Yaskawa INFORM job: VEGG2.JBI

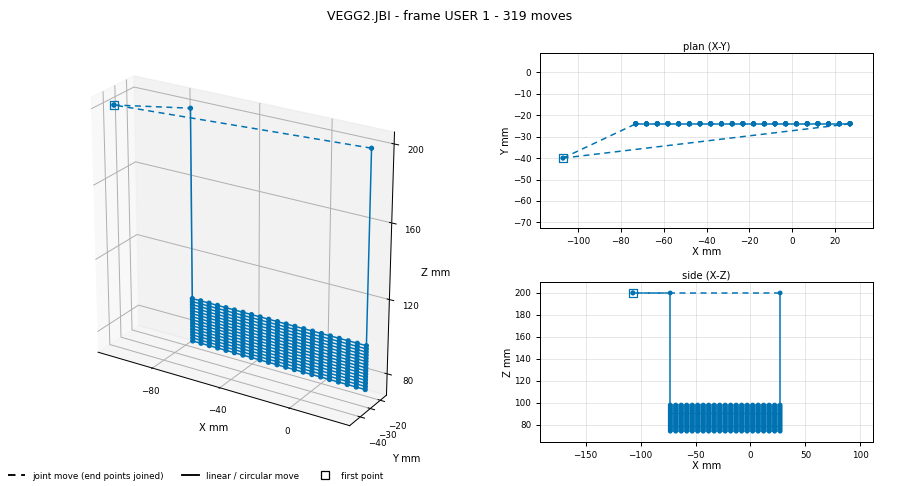
[picture p0: tool path of VEGG2.JBI in frame USER 1, 319 of 319 moves have a stored position in this frame; points joined in program order, loops and branches not executed]
/JOB
//NAME VEGG2
//POS
///NPOS 319,0,0,0,0,0
///USER 1
///TOOL 1
///POSTYPE USER
///RECTAN
///RCONF 1,0,0,0,0,0,0,0,0,0,0,0,0,0,0,0,0,0,0,0,0,0,0,0
C00000=-107.000,-40.000,200.000,0.0000,0.0000,-150.0000
C00001=-73.000,-24.000,200.000,0.0000,0.0000,-150.0000
C00002=-73.000,-24.000,74.200,0.0000,0.0000,-150.0000
C00003=-68.000,-24.000,74.200,0.0000,0.0000,-150.0000
C00004=-63.000,-24.000,74.200,0.0000,0.0000,-150.0000
C00005=-58.000,-24.000,74.200,0.0000,0.0000,-150.0000
C00006=-53.000,-24.000,74.200,0.0000,0.0000,-150.0000
C00007=-48.000,-24.000,74.200,0.0000,0.0000,-150.0000
C00008=-43.000,-24.000,74.200,0.0000,0.0000,-150.0000
C00009=-38.000,-24.000,74.200,0.0000,0.0000,-150.0000
C00010=-33.000,-24.000,74.200,0.0000,0.0000,-150.0000
C00011=-28.000,-24.000,74.200,0.0000,0.0000,-150.0000
C00012=-23.000,-24.000,74.200,0.0000,0.0000,-150.0000
C00013=-18.000,-24.000,74.200,0.0000,0.0000,-150.0000
C00014=-13.000,-24.000,74.200,0.0000,0.0000,-150.0000
C00015=-8.000,-24.000,74.200,0.0000,0.0000,-150.0000
C00016=-3.000,-24.000,74.200,0.0000,0.0000,-150.0000
C00017=2.000,-24.000,74.200,0.0000,0.0000,-150.0000
C00018=7.000,-24.000,74.200,0.0000,0.0000,-150.0000
C00019=12.000,-24.000,74.200,0.0000,0.0000,-150.0000
C00020=17.000,-24.000,74.200,0.0000,0.0000,-150.0000
C00021=22.000,-24.000,74.200,0.0000,0.0000,-150.0000
C00022=27.000,-24.000,74.200,0.0000,0.0000,-150.0000
C00023=27.000,-24.000,75.900,0.0000,0.0000,-150.0000
C00024=22.000,-24.000,75.900,0.0000,0.0000,-150.0000
C00025=17.000,-24.000,75.900,0.0000,0.0000,-150.0000
C00026=12.000,-24.000,75.900,0.0000,0.0000,-150.0000
C00027=7.000,-24.000,75.900,0.0000,0.0000,-150.0000
C00028=2.000,-24.000,75.900,0.0000,0.0000,-150.0000
C00029=-3.000,-24.000,75.900,0.0000,0.0000,-150.0000
C00030=-8.000,-24.000,75.900,0.0000,0.0000,-150.0000
C00031=-13.000,-24.000,75.900,0.0000,0.0000,-150.0000
C00032=-18.000,-24.000,75.900,0.0000,0.0000,-150.0000
C00033=-23.000,-24.000,75.900,0.0000,0.0000,-150.0000
C00034=-28.000,-24.000,75.900,0.0000,0.0000,-150.0000
C00035=-33.000,-24.000,75.900,0.0000,0.0000,-150.0000
C00036=-38.000,-24.000,75.900,0.0000,0.0000,-150.0000
C00037=-43.000,-24.000,75.900,0.0000,0.0000,-150.0000
C00038=-48.000,-24.000,75.900,0.0000,0.0000,-150.0000
C00039=-53.000,-24.000,75.900,0.0000,0.0000,-150.0000
C00040=-58.000,-24.000,75.900,0.0000,0.0000,-150.0000
C00041=-63.000,-24.000,75.900,0.0000,0.0000,-150.0000
C00042=-68.000,-24.000,75.900,0.0000,0.0000,-150.0000
C00043=-73.000,-24.000,75.900,0.0000,0.0000,-150.0000
C00044=-73.000,-24.000,77.600,0.0000,0.0000,-150.0000
C00045=-68.000,-24.000,77.600,0.0000,0.0000,-150.0000
C00046=-63.000,-24.000,77.600,0.0000,0.0000,-150.0000
C00047=-58.000,-24.000,77.600,0.0000,0.0000,-150.0000
C00048=-53.000,-24.000,77.600,0.0000,0.0000,-150.0000
C00049=-48.000,-24.000,77.600,0.0000,0.0000,-150.0000
C00050=-43.000,-24.000,77.600,0.0000,0.0000,-150.0000
C00051=-38.000,-24.000,77.600,0.0000,0.0000,-150.0000
C00052=-33.000,-24.000,77.600,0.0000,0.0000,-150.0000
C00053=-28.000,-24.000,77.600,0.0000,0.0000,-150.0000
C00054=-23.000,-24.000,77.600,0.0000,0.0000,-150.0000
C00055=-18.000,-24.000,77.600,0.0000,0.0000,-150.0000
C00056=-13.000,-24.000,77.600,0.0000,0.0000,-150.0000
C00057=-8.000,-24.000,77.600,0.0000,0.0000,-150.0000
C00058=-3.000,-24.000,77.600,0.0000,0.0000,-150.0000
C00059=2.000,-24.000,77.600,0.0000,0.0000,-150.0000
C00060=7.000,-24.000,77.600,0.0000,0.0000,-150.0000
C00061=12.000,-24.000,77.600,0.0000,0.0000,-150.0000
C00062=17.000,-24.000,77.600,0.0000,0.0000,-150.0000
C00063=22.000,-24.000,77.600,0.0000,0.0000,-150.0000
C00064=27.000,-24.000,77.600,0.0000,0.0000,-150.0000
C00065=27.000,-24.000,79.300,0.0000,0.0000,-150.0000
C00066=22.000,-24.000,79.300,0.0000,0.0000,-150.0000
C00067=17.000,-24.000,79.300,0.0000,0.0000,-150.0000
C00068=12.000,-24.000,79.300,0.0000,0.0000,-150.0000
C00069=7.000,-24.000,79.300,0.0000,0.0000,-150.0000
C00070=2.000,-24.000,79.300,0.0000,0.0000,-150.0000
C00071=-3.000,-24.000,79.300,0.0000,0.0000,-150.0000
C00072=-8.000,-24.000,79.300,0.0000,0.0000,-150.0000
C00073=-13.000,-24.000,79.300,0.0000,0.0000,-150.0000
C00074=-18.000,-24.000,79.300,0.0000,0.0000,-150.0000
C00075=-23.000,-24.000,79.300,0.0000,0.0000,-150.0000
C00076=-28.000,-24.000,79.300,0.0000,0.0000,-150.0000
C00077=-33.000,-24.000,79.300,0.0000,0.0000,-150.0000
C00078=-38.000,-24.000,79.300,0.0000,0.0000,-150.0000
C00079=-43.000,-24.000,79.300,0.0000,0.0000,-150.0000
C00080=-48.000,-24.000,79.300,0.0000,0.0000,-150.0000
C00081=-53.000,-24.000,79.300,0.0000,0.0000,-150.0000
C00082=-58.000,-24.000,79.300,0.0000,0.0000,-150.0000
C00083=-63.000,-24.000,79.300,0.0000,0.0000,-150.0000
C00084=-68.000,-24.000,79.300,0.0000,0.0000,-150.0000
C00085=-73.000,-24.000,79.300,0.0000,0.0000,-150.0000
C00086=-73.000,-24.000,81.000,0.0000,0.0000,-150.0000
C00087=-68.000,-24.000,81.000,0.0000,0.0000,-150.0000
C00088=-63.000,-24.000,81.000,0.0000,0.0000,-150.0000
C00089=-58.000,-24.000,81.000,0.0000,0.0000,-150.0000
C00090=-53.000,-24.000,81.000,0.0000,0.0000,-150.0000
C00091=-48.000,-24.000,81.000,0.0000,0.0000,-150.0000
C00092=-43.000,-24.000,81.000,0.0000,0.0000,-150.0000
C00093=-38.000,-24.000,81.000,0.0000,0.0000,-150.0000
C00094=-33.000,-24.000,81.000,0.0000,0.0000,-150.0000
C00095=-28.000,-24.000,81.000,0.0000,0.0000,-150.0000
C00096=-23.000,-24.000,81.000,0.0000,0.0000,-150.0000
C00097=-18.000,-24.000,81.000,0.0000,0.0000,-150.0000
C00098=-13.000,-24.000,81.000,0.0000,0.0000,-150.0000
C00099=-8.000,-24.000,81.000,0.0000,0.0000,-150.0000
C00100=-3.000,-24.000,81.000,0.0000,0.0000,-150.0000
C00101=2.000,-24.000,81.000,0.0000,0.0000,-150.0000
C00102=7.000,-24.000,81.000,0.0000,0.0000,-150.0000
C00103=12.000,-24.000,81.000,0.0000,0.0000,-150.0000
C00104=17.000,-24.000,81.000,0.0000,0.0000,-150.0000
C00105=22.000,-24.000,81.000,0.0000,0.0000,-150.0000
C00106=27.000,-24.000,81.000,0.0000,0.0000,-150.0000
C00107=27.000,-24.000,82.700,0.0000,0.0000,-150.0000
C00108=22.000,-24.000,82.700,0.0000,0.0000,-150.0000
C00109=17.000,-24.000,82.700,0.0000,0.0000,-150.0000
C00110=12.000,-24.000,82.700,0.0000,0.0000,-150.0000
C00111=7.000,-24.000,82.700,0.0000,0.0000,-150.0000
C00112=2.000,-24.000,82.700,0.0000,0.0000,-150.0000
C00113=-3.000,-24.000,82.700,0.0000,0.0000,-150.0000
C00114=-8.000,-24.000,82.700,0.0000,0.0000,-150.0000
C00115=-13.000,-24.000,82.700,0.0000,0.0000,-150.0000
C00116=-18.000,-24.000,82.700,0.0000,0.0000,-150.0000
C00117=-23.000,-24.000,82.700,0.0000,0.0000,-150.0000
C00118=-28.000,-24.000,82.700,0.0000,0.0000,-150.0000
C00119=-33.000,-24.000,82.700,0.0000,0.0000,-150.0000
C00120=-38.000,-24.000,82.700,0.0000,0.0000,-150.0000
C00121=-43.000,-24.000,82.700,0.0000,0.0000,-150.0000
C00122=-48.000,-24.000,82.700,0.0000,0.0000,-150.0000
C00123=-53.000,-24.000,82.700,0.0000,0.0000,-150.0000
C00124=-58.000,-24.000,82.700,0.0000,0.0000,-150.0000
C00125=-63.000,-24.000,82.700,0.0000,0.0000,-150.0000
C00126=-68.000,-24.000,82.700,0.0000,0.0000,-150.0000
C00127=-73.000,-24.000,82.700,0.0000,0.0000,-150.0000
C00128=-73.000,-24.000,84.400,0.0000,0.0000,-150.0000
C00129=-68.000,-24.000,84.400,0.0000,0.0000,-150.0000
C00130=-63.000,-24.000,84.400,0.0000,0.0000,-150.0000
C00131=-58.000,-24.000,84.400,0.0000,0.0000,-150.0000
C00132=-53.000,-24.000,84.400,0.0000,0.0000,-150.0000
C00133=-48.000,-24.000,84.400,0.0000,0.0000,-150.0000
C00134=-43.000,-24.000,84.400,0.0000,0.0000,-150.0000
C00135=-38.000,-24.000,84.400,0.0000,0.0000,-150.0000
C00136=-33.000,-24.000,84.400,0.0000,0.0000,-150.0000
C00137=-28.000,-24.000,84.400,0.0000,0.0000,-150.0000
C00138=-23.000,-24.000,84.400,0.0000,0.0000,-150.0000
C00139=-18.000,-24.000,84.400,0.0000,0.0000,-150.0000
C00140=-13.000,-24.000,84.400,0.0000,0.0000,-150.0000
C00141=-8.000,-24.000,84.400,0.0000,0.0000,-150.0000
C00142=-3.000,-24.000,84.400,0.0000,0.0000,-150.0000
C00143=2.000,-24.000,84.400,0.0000,0.0000,-150.0000
C00144=7.000,-24.000,84.400,0.0000,0.0000,-150.0000
C00145=12.000,-24.000,84.400,0.0000,0.0000,-150.0000
C00146=17.000,-24.000,84.400,0.0000,0.0000,-150.0000
C00147=22.000,-24.000,84.400,0.0000,0.0000,-150.0000
C00148=27.000,-24.000,84.400,0.0000,0.0000,-150.0000
C00149=27.000,-24.000,86.100,0.0000,0.0000,-150.0000
C00150=22.000,-24.000,86.100,0.0000,0.0000,-150.0000
C00151=17.000,-24.000,86.100,0.0000,0.0000,-150.0000
C00152=12.000,-24.000,86.100,0.0000,0.0000,-150.0000
C00153=7.000,-24.000,86.100,0.0000,0.0000,-150.0000
C00154=2.000,-24.000,86.100,0.0000,0.0000,-150.0000
C00155=-3.000,-24.000,86.100,0.0000,0.0000,-150.0000
C00156=-8.000,-24.000,86.100,0.0000,0.0000,-150.0000
C00157=-13.000,-24.000,86.100,0.0000,0.0000,-150.0000
C00158=-18.000,-24.000,86.100,0.0000,0.0000,-150.0000
C00159=-23.000,-24.000,86.100,0.0000,0.0000,-150.0000
C00160=-28.000,-24.000,86.100,0.0000,0.0000,-150.0000
C00161=-33.000,-24.000,86.100,0.0000,0.0000,-150.0000
C00162=-38.000,-24.000,86.100,0.0000,0.0000,-150.0000
C00163=-43.000,-24.000,86.100,0.0000,0.0000,-150.0000
C00164=-48.000,-24.000,86.100,0.0000,0.0000,-150.0000
C00165=-53.000,-24.000,86.100,0.0000,0.0000,-150.0000
C00166=-58.000,-24.000,86.100,0.0000,0.0000,-150.0000
C00167=-63.000,-24.000,86.100,0.0000,0.0000,-150.0000
C00168=-68.000,-24.000,86.100,0.0000,0.0000,-150.0000
C00169=-73.000,-24.000,86.100,0.0000,0.0000,-150.0000
C00170=-73.000,-24.000,87.800,0.0000,0.0000,-150.0000
C00171=-68.000,-24.000,87.800,0.0000,0.0000,-150.0000
C00172=-63.000,-24.000,87.800,0.0000,0.0000,-150.0000
C00173=-58.000,-24.000,87.800,0.0000,0.0000,-150.0000
C00174=-53.000,-24.000,87.800,0.0000,0.0000,-150.0000
C00175=-48.000,-24.000,87.800,0.0000,0.0000,-150.0000
C00176=-43.000,-24.000,87.800,0.0000,0.0000,-150.0000
C00177=-38.000,-24.000,87.800,0.0000,0.0000,-150.0000
C00178=-33.000,-24.000,87.800,0.0000,0.0000,-150.0000
C00179=-28.000,-24.000,87.800,0.0000,0.0000,-150.0000
C00180=-23.000,-24.000,87.800,0.0000,0.0000,-150.0000
C00181=-18.000,-24.000,87.800,0.0000,0.0000,-150.0000
C00182=-13.000,-24.000,87.800,0.0000,0.0000,-150.0000
C00183=-8.000,-24.000,87.800,0.0000,0.0000,-150.0000
C00184=-3.000,-24.000,87.800,0.0000,0.0000,-150.0000
C00185=2.000,-24.000,87.800,0.0000,0.0000,-150.0000
C00186=7.000,-24.000,87.800,0.0000,0.0000,-150.0000
C00187=12.000,-24.000,87.800,0.0000,0.0000,-150.0000
C00188=17.000,-24.000,87.800,0.0000,0.0000,-150.0000
C00189=22.000,-24.000,87.800,0.0000,0.0000,-150.0000
C00190=27.000,-24.000,87.800,0.0000,0.0000,-150.0000
C00191=27.000,-24.000,89.500,0.0000,0.0000,-150.0000
C00192=22.000,-24.000,89.500,0.0000,0.0000,-150.0000
C00193=17.000,-24.000,89.500,0.0000,0.0000,-150.0000
C00194=12.000,-24.000,89.500,0.0000,0.0000,-150.0000
C00195=7.000,-24.000,89.500,0.0000,0.0000,-150.0000
C00196=2.000,-24.000,89.500,0.0000,0.0000,-150.0000
C00197=-3.000,-24.000,89.500,0.0000,0.0000,-150.0000
C00198=-8.000,-24.000,89.500,0.0000,0.0000,-150.0000
C00199=-13.000,-24.000,89.500,0.0000,0.0000,-150.0000
C00200=-18.000,-24.000,89.500,0.0000,0.0000,-150.0000
C00201=-23.000,-24.000,89.500,0.0000,0.0000,-150.0000
C00202=-28.000,-24.000,89.500,0.0000,0.0000,-150.0000
C00203=-33.000,-24.000,89.500,0.0000,0.0000,-150.0000
C00204=-38.000,-24.000,89.500,0.0000,0.0000,-150.0000
C00205=-43.000,-24.000,89.500,0.0000,0.0000,-150.0000
C00206=-48.000,-24.000,89.500,0.0000,0.0000,-150.0000
C00207=-53.000,-24.000,89.500,0.0000,0.0000,-150.0000
C00208=-58.000,-24.000,89.500,0.0000,0.0000,-150.0000
C00209=-63.000,-24.000,89.500,0.0000,0.0000,-150.0000
C00210=-68.000,-24.000,89.500,0.0000,0.0000,-150.0000
C00211=-73.000,-24.000,89.500,0.0000,0.0000,-150.0000
C00212=-73.000,-24.000,91.200,0.0000,0.0000,-150.0000
C00213=-68.000,-24.000,91.200,0.0000,0.0000,-150.0000
C00214=-63.000,-24.000,91.200,0.0000,0.0000,-150.0000
C00215=-58.000,-24.000,91.200,0.0000,0.0000,-150.0000
C00216=-53.000,-24.000,91.200,0.0000,0.0000,-150.0000
C00217=-48.000,-24.000,91.200,0.0000,0.0000,-150.0000
C00218=-43.000,-24.000,91.200,0.0000,0.0000,-150.0000
C00219=-38.000,-24.000,91.200,0.0000,0.0000,-150.0000
C00220=-33.000,-24.000,91.200,0.0000,0.0000,-150.0000
C00221=-28.000,-24.000,91.200,0.0000,0.0000,-150.0000
C00222=-23.000,-24.000,91.200,0.0000,0.0000,-150.0000
C00223=-18.000,-24.000,91.200,0.0000,0.0000,-150.0000
C00224=-13.000,-24.000,91.200,0.0000,0.0000,-150.0000
C00225=-8.000,-24.000,91.200,0.0000,0.0000,-150.0000
C00226=-3.000,-24.000,91.200,0.0000,0.0000,-150.0000
C00227=2.000,-24.000,91.200,0.0000,0.0000,-150.0000
C00228=7.000,-24.000,91.200,0.0000,0.0000,-150.0000
C00229=12.000,-24.000,91.200,0.0000,0.0000,-150.0000
C00230=17.000,-24.000,91.200,0.0000,0.0000,-150.0000
C00231=22.000,-24.000,91.200,0.0000,0.0000,-150.0000
C00232=27.000,-24.000,91.200,0.0000,0.0000,-150.0000
C00233=27.000,-24.000,92.900,0.0000,0.0000,-150.0000
C00234=22.000,-24.000,92.900,0.0000,0.0000,-150.0000
C00235=17.000,-24.000,92.900,0.0000,0.0000,-150.0000
C00236=12.000,-24.000,92.900,0.0000,0.0000,-150.0000
C00237=7.000,-24.000,92.900,0.0000,0.0000,-150.0000
C00238=2.000,-24.000,92.900,0.0000,0.0000,-150.0000
C00239=-3.000,-24.000,92.900,0.0000,0.0000,-150.0000
C00240=-8.000,-24.000,92.900,0.0000,0.0000,-150.0000
C00241=-13.000,-24.000,92.900,0.0000,0.0000,-150.0000
C00242=-18.000,-24.000,92.900,0.0000,0.0000,-150.0000
C00243=-23.000,-24.000,92.900,0.0000,0.0000,-150.0000
C00244=-28.000,-24.000,92.900,0.0000,0.0000,-150.0000
C00245=-33.000,-24.000,92.900,0.0000,0.0000,-150.0000
C00246=-38.000,-24.000,92.900,0.0000,0.0000,-150.0000
C00247=-43.000,-24.000,92.900,0.0000,0.0000,-150.0000
C00248=-48.000,-24.000,92.900,0.0000,0.0000,-150.0000
C00249=-53.000,-24.000,92.900,0.0000,0.0000,-150.0000
C00250=-58.000,-24.000,92.900,0.0000,0.0000,-150.0000
C00251=-63.000,-24.000,92.900,0.0000,0.0000,-150.0000
C00252=-68.000,-24.000,92.900,0.0000,0.0000,-150.0000
C00253=-73.000,-24.000,92.900,0.0000,0.0000,-150.0000
C00254=-73.000,-24.000,94.600,0.0000,0.0000,-150.0000
C00255=-68.000,-24.000,94.600,0.0000,0.0000,-150.0000
C00256=-63.000,-24.000,94.600,0.0000,0.0000,-150.0000
C00257=-58.000,-24.000,94.600,0.0000,0.0000,-150.0000
C00258=-53.000,-24.000,94.600,0.0000,0.0000,-150.0000
C00259=-48.000,-24.000,94.600,0.0000,0.0000,-150.0000
C00260=-43.000,-24.000,94.600,0.0000,0.0000,-150.0000
C00261=-38.000,-24.000,94.600,0.0000,0.0000,-150.0000
C00262=-33.000,-24.000,94.600,0.0000,0.0000,-150.0000
C00263=-28.000,-24.000,94.600,0.0000,0.0000,-150.0000
C00264=-23.000,-24.000,94.600,0.0000,0.0000,-150.0000
C00265=-18.000,-24.000,94.600,0.0000,0.0000,-150.0000
C00266=-13.000,-24.000,94.600,0.0000,0.0000,-150.0000
C00267=-8.000,-24.000,94.600,0.0000,0.0000,-150.0000
C00268=-3.000,-24.000,94.600,0.0000,0.0000,-150.0000
C00269=2.000,-24.000,94.600,0.0000,0.0000,-150.0000
C00270=7.000,-24.000,94.600,0.0000,0.0000,-150.0000
C00271=12.000,-24.000,94.600,0.0000,0.0000,-150.0000
C00272=17.000,-24.000,94.600,0.0000,0.0000,-150.0000
C00273=22.000,-24.000,94.600,0.0000,0.0000,-150.0000
C00274=27.000,-24.000,94.600,0.0000,0.0000,-150.0000
C00275=27.000,-24.000,96.300,0.0000,0.0000,-150.0000
C00276=22.000,-24.000,96.300,0.0000,0.0000,-150.0000
C00277=17.000,-24.000,96.300,0.0000,0.0000,-150.0000
C00278=12.000,-24.000,96.300,0.0000,0.0000,-150.0000
C00279=7.000,-24.000,96.300,0.0000,0.0000,-150.0000
C00280=2.000,-24.000,96.300,0.0000,0.0000,-150.0000
C00281=-3.000,-24.000,96.300,0.0000,0.0000,-150.0000
C00282=-8.000,-24.000,96.300,0.0000,0.0000,-150.0000
C00283=-13.000,-24.000,96.300,0.0000,0.0000,-150.0000
C00284=-18.000,-24.000,96.300,0.0000,0.0000,-150.0000
C00285=-23.000,-24.000,96.300,0.0000,0.0000,-150.0000
C00286=-28.000,-24.000,96.300,0.0000,0.0000,-150.0000
C00287=-33.000,-24.000,96.300,0.0000,0.0000,-150.0000
C00288=-38.000,-24.000,96.300,0.0000,0.0000,-150.0000
C00289=-43.000,-24.000,96.300,0.0000,0.0000,-150.0000
C00290=-48.000,-24.000,96.300,0.0000,0.0000,-150.0000
C00291=-53.000,-24.000,96.300,0.0000,0.0000,-150.0000
C00292=-58.000,-24.000,96.300,0.0000,0.0000,-150.0000
C00293=-63.000,-24.000,96.300,0.0000,0.0000,-150.0000
C00294=-68.000,-24.000,96.300,0.0000,0.0000,-150.0000
C00295=-73.000,-24.000,96.300,0.0000,0.0000,-150.0000
C00296=-73.000,-24.000,98.000,0.0000,0.0000,-150.0000
C00297=-68.000,-24.000,98.000,0.0000,0.0000,-150.0000
C00298=-63.000,-24.000,98.000,0.0000,0.0000,-150.0000
C00299=-58.000,-24.000,98.000,0.0000,0.0000,-150.0000
C00300=-53.000,-24.000,98.000,0.0000,0.0000,-150.0000
C00301=-48.000,-24.000,98.000,0.0000,0.0000,-150.0000
C00302=-43.000,-24.000,98.000,0.0000,0.0000,-150.0000
C00303=-38.000,-24.000,98.000,0.0000,0.0000,-150.0000
C00304=-33.000,-24.000,98.000,0.0000,0.0000,-150.0000
C00305=-28.000,-24.000,98.000,0.0000,0.0000,-150.0000
C00306=-23.000,-24.000,98.000,0.0000,0.0000,-150.0000
C00307=-18.000,-24.000,98.000,0.0000,0.0000,-150.0000
C00308=-13.000,-24.000,98.000,0.0000,0.0000,-150.0000
C00309=-8.000,-24.000,98.000,0.0000,0.0000,-150.0000
C00310=-3.000,-24.000,98.000,0.0000,0.0000,-150.0000
C00311=2.000,-24.000,98.000,0.0000,0.0000,-150.0000
C00312=7.000,-24.000,98.000,0.0000,0.0000,-150.0000
C00313=12.000,-24.000,98.000,0.0000,0.0000,-150.0000
C00314=17.000,-24.000,98.000,0.0000,0.0000,-150.0000
C00315=22.000,-24.000,98.000,0.0000,0.0000,-150.0000
C00316=27.000,-24.000,98.000,0.0000,0.0000,-150.0000
C00317=27.000,-24.000,200.000,0.0000,0.0000,-150.0000
C00318=-107.000,-40.000,200.000,0.0000,0.0000,-150.0000
//INST
///DATE 2026/11/20 16:20
///ATTR SC,RW,RJ
////FRAME USER 1
///GROUP1 RB1
NOP
MOVJ C00000 VJ=0.78
MOVJ C00001 VJ=0.78
MOVL C00002 V=7.0 ACC=20 DEC=20
*LAG1
MACRO1 MJ#(0) ARGF1
ARCON
MOVL C00003 V=7.0 ACC=20 DEC=20
MOVL C00004 V=7.0 ACC=20 DEC=20
MOVL C00005 V=7.0 ACC=20 DEC=20
MOVL C00006 V=7.0 ACC=20 DEC=20
MOVL C00007 V=7.0 ACC=20 DEC=20
MOVL C00008 V=7.0 ACC=20 DEC=20
MOVL C00009 V=7.0 ACC=20 DEC=20
MOVL C00010 V=7.0 ACC=20 DEC=20
MOVL C00011 V=7.0 ACC=20 DEC=20
MOVL C00012 V=7.0 ACC=20 DEC=20
MOVL C00013 V=7.0 ACC=20 DEC=20
MOVL C00014 V=7.0 ACC=20 DEC=20
MOVL C00015 V=7.0 ACC=20 DEC=20
MOVL C00016 V=7.0 ACC=20 DEC=20
MOVL C00017 V=7.0 ACC=20 DEC=20
MOVL C00018 V=7.0 ACC=20 DEC=20
MOVL C00019 V=7.0 ACC=20 DEC=20
MOVL C00020 V=7.0 ACC=20 DEC=20
MOVL C00021 V=7.0 ACC=20 DEC=20
MOVL C00022 V=7.0 ACC=20 DEC=20
ARCOF
TIMER T=30
*LAG2
MOVL C00023 V=7.0 ACC=20 DEC=20
MACRO1 MJ#(0) ARGF2
ARCON
MOVL C00024 V=7.0 ACC=20 DEC=20
MOVL C00025 V=7.0 ACC=20 DEC=20
MOVL C00026 V=7.0 ACC=20 DEC=20
MOVL C00027 V=7.0 ACC=20 DEC=20
MOVL C00028 V=7.0 ACC=20 DEC=20
MOVL C00029 V=7.0 ACC=20 DEC=20
MOVL C00030 V=7.0 ACC=20 DEC=20
MOVL C00031 V=7.0 ACC=20 DEC=20
MOVL C00032 V=7.0 ACC=20 DEC=20
MOVL C00033 V=7.0 ACC=20 DEC=20
MOVL C00034 V=7.0 ACC=20 DEC=20
MOVL C00035 V=7.0 ACC=20 DEC=20
MOVL C00036 V=7.0 ACC=20 DEC=20
MOVL C00037 V=7.0 ACC=20 DEC=20
MOVL C00038 V=7.0 ACC=20 DEC=20
MOVL C00039 V=7.0 ACC=20 DEC=20
MOVL C00040 V=7.0 ACC=20 DEC=20
MOVL C00041 V=7.0 ACC=20 DEC=20
MOVL C00042 V=7.0 ACC=20 DEC=20
MOVL C00043 V=7.0 ACC=20 DEC=20
ARCOF
TIMER T=30
*LAG3
MOVL C00044 V=7.0 ACC=20 DEC=20
MACRO1 MJ#(0) ARGF2
ARCON
MOVL C00045 V=7.0 ACC=20 DEC=20
MOVL C00046 V=7.0 ACC=20 DEC=20
MOVL C00047 V=7.0 ACC=20 DEC=20
MOVL C00048 V=7.0 ACC=20 DEC=20
MOVL C00049 V=7.0 ACC=20 DEC=20
MOVL C00050 V=7.0 ACC=20 DEC=20
MOVL C00051 V=7.0 ACC=20 DEC=20
MOVL C00052 V=7.0 ACC=20 DEC=20
MOVL C00053 V=7.0 ACC=20 DEC=20
MOVL C00054 V=7.0 ACC=20 DEC=20
MOVL C00055 V=7.0 ACC=20 DEC=20
MOVL C00056 V=7.0 ACC=20 DEC=20
MOVL C00057 V=7.0 ACC=20 DEC=20
MOVL C00058 V=7.0 ACC=20 DEC=20
MOVL C00059 V=7.0 ACC=20 DEC=20
MOVL C00060 V=7.0 ACC=20 DEC=20
MOVL C00061 V=7.0 ACC=20 DEC=20
MOVL C00062 V=7.0 ACC=20 DEC=20
MOVL C00063 V=7.0 ACC=20 DEC=20
MOVL C00064 V=7.0 ACC=20 DEC=20
ARCOF
TIMER T=30
*LAG4
MOVL C00065 V=7.0 ACC=20 DEC=20
MACRO1 MJ#(0) ARGF2
ARCON
MOVL C00066 V=7.0 ACC=20 DEC=20
MOVL C00067 V=7.0 ACC=20 DEC=20
MOVL C00068 V=7.0 ACC=20 DEC=20
MOVL C00069 V=7.0 ACC=20 DEC=20
MOVL C00070 V=7.0 ACC=20 DEC=20
MOVL C00071 V=7.0 ACC=20 DEC=20
MOVL C00072 V=7.0 ACC=20 DEC=20
MOVL C00073 V=7.0 ACC=20 DEC=20
MOVL C00074 V=7.0 ACC=20 DEC=20
MOVL C00075 V=7.0 ACC=20 DEC=20
MOVL C00076 V=7.0 ACC=20 DEC=20
MOVL C00077 V=7.0 ACC=20 DEC=20
MOVL C00078 V=7.0 ACC=20 DEC=20
MOVL C00079 V=7.0 ACC=20 DEC=20
MOVL C00080 V=7.0 ACC=20 DEC=20
MOVL C00081 V=7.0 ACC=20 DEC=20
MOVL C00082 V=7.0 ACC=20 DEC=20
MOVL C00083 V=7.0 ACC=20 DEC=20
MOVL C00084 V=7.0 ACC=20 DEC=20
MOVL C00085 V=7.0 ACC=20 DEC=20
ARCOF
TIMER T=30
*LAG5
MOVL C00086 V=7.0 ACC=20 DEC=20
MACRO1 MJ#(0) ARGF2
ARCON
MOVL C00087 V=7.0 ACC=20 DEC=20
MOVL C00088 V=7.0 ACC=20 DEC=20
MOVL C00089 V=7.0 ACC=20 DEC=20
MOVL C00090 V=7.0 ACC=20 DEC=20
MOVL C00091 V=7.0 ACC=20 DEC=20
MOVL C00092 V=7.0 ACC=20 DEC=20
MOVL C00093 V=7.0 ACC=20 DEC=20
MOVL C00094 V=7.0 ACC=20 DEC=20
MOVL C00095 V=7.0 ACC=20 DEC=20
MOVL C00096 V=7.0 ACC=20 DEC=20
MOVL C00097 V=7.0 ACC=20 DEC=20
MOVL C00098 V=7.0 ACC=20 DEC=20
MOVL C00099 V=7.0 ACC=20 DEC=20
MOVL C00100 V=7.0 ACC=20 DEC=20
MOVL C00101 V=7.0 ACC=20 DEC=20
MOVL C00102 V=7.0 ACC=20 DEC=20
MOVL C00103 V=7.0 ACC=20 DEC=20
MOVL C00104 V=7.0 ACC=20 DEC=20
MOVL C00105 V=7.0 ACC=20 DEC=20
MOVL C00106 V=7.0 ACC=20 DEC=20
ARCOF
TIMER T=30
*LAG6
MOVL C00107 V=7.0 ACC=20 DEC=20
MACRO1 MJ#(0) ARGF2
ARCON
MOVL C00108 V=7.0 ACC=20 DEC=20
MOVL C00109 V=7.0 ACC=20 DEC=20
MOVL C00110 V=7.0 ACC=20 DEC=20
MOVL C00111 V=7.0 ACC=20 DEC=20
MOVL C00112 V=7.0 ACC=20 DEC=20
MOVL C00113 V=7.0 ACC=20 DEC=20
MOVL C00114 V=7.0 ACC=20 DEC=20
MOVL C00115 V=7.0 ACC=20 DEC=20
MOVL C00116 V=7.0 ACC=20 DEC=20
MOVL C00117 V=7.0 ACC=20 DEC=20
MOVL C00118 V=7.0 ACC=20 DEC=20
MOVL C00119 V=7.0 ACC=20 DEC=20
MOVL C00120 V=7.0 ACC=20 DEC=20
MOVL C00121 V=7.0 ACC=20 DEC=20
MOVL C00122 V=7.0 ACC=20 DEC=20
MOVL C00123 V=7.0 ACC=20 DEC=20
MOVL C00124 V=7.0 ACC=20 DEC=20
MOVL C00125 V=7.0 ACC=20 DEC=20
MOVL C00126 V=7.0 ACC=20 DEC=20
MOVL C00127 V=7.0 ACC=20 DEC=20
ARCOF
TIMER T=30
*LAG7
MOVL C00128 V=7.0 ACC=20 DEC=20
MACRO1 MJ#(0) ARGF2
ARCON
MOVL C00129 V=7.0 ACC=20 DEC=20
MOVL C00130 V=7.0 ACC=20 DEC=20
MOVL C00131 V=7.0 ACC=20 DEC=20
MOVL C00132 V=7.0 ACC=20 DEC=20
MOVL C00133 V=7.0 ACC=20 DEC=20
MOVL C00134 V=7.0 ACC=20 DEC=20
MOVL C00135 V=7.0 ACC=20 DEC=20
MOVL C00136 V=7.0 ACC=20 DEC=20
MOVL C00137 V=7.0 ACC=20 DEC=20
MOVL C00138 V=7.0 ACC=20 DEC=20
MOVL C00139 V=7.0 ACC=20 DEC=20
MOVL C00140 V=7.0 ACC=20 DEC=20
MOVL C00141 V=7.0 ACC=20 DEC=20
MOVL C00142 V=7.0 ACC=20 DEC=20
MOVL C00143 V=7.0 ACC=20 DEC=20
MOVL C00144 V=7.0 ACC=20 DEC=20
MOVL C00145 V=7.0 ACC=20 DEC=20
MOVL C00146 V=7.0 ACC=20 DEC=20
MOVL C00147 V=7.0 ACC=20 DEC=20
MOVL C00148 V=7.0 ACC=20 DEC=20
ARCOF
TIMER T=30
*LAG8
MOVL C00149 V=7.0 ACC=20 DEC=20
MACRO1 MJ#(0) ARGF2
ARCON
MOVL C00150 V=7.0 ACC=20 DEC=20
MOVL C00151 V=7.0 ACC=20 DEC=20
MOVL C00152 V=7.0 ACC=20 DEC=20
MOVL C00153 V=7.0 ACC=20 DEC=20
MOVL C00154 V=7.0 ACC=20 DEC=20
MOVL C00155 V=7.0 ACC=20 DEC=20
MOVL C00156 V=7.0 ACC=20 DEC=20
MOVL C00157 V=7.0 ACC=20 DEC=20
MOVL C00158 V=7.0 ACC=20 DEC=20
MOVL C00159 V=7.0 ACC=20 DEC=20
MOVL C00160 V=7.0 ACC=20 DEC=20
MOVL C00161 V=7.0 ACC=20 DEC=20
MOVL C00162 V=7.0 ACC=20 DEC=20
MOVL C00163 V=7.0 ACC=20 DEC=20
MOVL C00164 V=7.0 ACC=20 DEC=20
MOVL C00165 V=7.0 ACC=20 DEC=20
MOVL C00166 V=7.0 ACC=20 DEC=20
MOVL C00167 V=7.0 ACC=20 DEC=20
MOVL C00168 V=7.0 ACC=20 DEC=20
MOVL C00169 V=7.0 ACC=20 DEC=20
ARCOF
TIMER T=30
*LAG9
MOVL C00170 V=7.0 ACC=20 DEC=20
MACRO1 MJ#(0) ARGF2
ARCON
MOVL C00171 V=7.0 ACC=20 DEC=20
MOVL C00172 V=7.0 ACC=20 DEC=20
MOVL C00173 V=7.0 ACC=20 DEC=20
MOVL C00174 V=7.0 ACC=20 DEC=20
MOVL C00175 V=7.0 ACC=20 DEC=20
MOVL C00176 V=7.0 ACC=20 DEC=20
MOVL C00177 V=7.0 ACC=20 DEC=20
MOVL C00178 V=7.0 ACC=20 DEC=20
MOVL C00179 V=7.0 ACC=20 DEC=20
MOVL C00180 V=7.0 ACC=20 DEC=20
MOVL C00181 V=7.0 ACC=20 DEC=20
MOVL C00182 V=7.0 ACC=20 DEC=20
MOVL C00183 V=7.0 ACC=20 DEC=20
MOVL C00184 V=7.0 ACC=20 DEC=20
MOVL C00185 V=7.0 ACC=20 DEC=20
MOVL C00186 V=7.0 ACC=20 DEC=20
MOVL C00187 V=7.0 ACC=20 DEC=20
MOVL C00188 V=7.0 ACC=20 DEC=20
MOVL C00189 V=7.0 ACC=20 DEC=20
MOVL C00190 V=7.0 ACC=20 DEC=20
ARCOF
TIMER T=30
*LAG10
MOVL C00191 V=7.0 ACC=20 DEC=20
MACRO1 MJ#(0) ARGF2
ARCON
MOVL C00192 V=7.0 ACC=20 DEC=20
MOVL C00193 V=7.0 ACC=20 DEC=20
MOVL C00194 V=7.0 ACC=20 DEC=20
MOVL C00195 V=7.0 ACC=20 DEC=20
MOVL C00196 V=7.0 ACC=20 DEC=20
MOVL C00197 V=7.0 ACC=20 DEC=20
MOVL C00198 V=7.0 ACC=20 DEC=20
MOVL C00199 V=7.0 ACC=20 DEC=20
MOVL C00200 V=7.0 ACC=20 DEC=20
MOVL C00201 V=7.0 ACC=20 DEC=20
MOVL C00202 V=7.0 ACC=20 DEC=20
MOVL C00203 V=7.0 ACC=20 DEC=20
MOVL C00204 V=7.0 ACC=20 DEC=20
MOVL C00205 V=7.0 ACC=20 DEC=20
MOVL C00206 V=7.0 ACC=20 DEC=20
MOVL C00207 V=7.0 ACC=20 DEC=20
MOVL C00208 V=7.0 ACC=20 DEC=20
MOVL C00209 V=7.0 ACC=20 DEC=20
MOVL C00210 V=7.0 ACC=20 DEC=20
MOVL C00211 V=7.0 ACC=20 DEC=20
ARCOF
TIMER T=30
*LAG11
MOVL C00212 V=7.0 ACC=20 DEC=20
MACRO1 MJ#(0) ARGF2
ARCON
MOVL C00213 V=7.0 ACC=20 DEC=20
MOVL C00214 V=7.0 ACC=20 DEC=20
MOVL C00215 V=7.0 ACC=20 DEC=20
MOVL C00216 V=7.0 ACC=20 DEC=20
MOVL C00217 V=7.0 ACC=20 DEC=20
MOVL C00218 V=7.0 ACC=20 DEC=20
MOVL C00219 V=7.0 ACC=20 DEC=20
MOVL C00220 V=7.0 ACC=20 DEC=20
MOVL C00221 V=7.0 ACC=20 DEC=20
MOVL C00222 V=7.0 ACC=20 DEC=20
MOVL C00223 V=7.0 ACC=20 DEC=20
MOVL C00224 V=7.0 ACC=20 DEC=20
MOVL C00225 V=7.0 ACC=20 DEC=20
MOVL C00226 V=7.0 ACC=20 DEC=20
MOVL C00227 V=7.0 ACC=20 DEC=20
MOVL C00228 V=7.0 ACC=20 DEC=20
MOVL C00229 V=7.0 ACC=20 DEC=20
MOVL C00230 V=7.0 ACC=20 DEC=20
MOVL C00231 V=7.0 ACC=20 DEC=20
MOVL C00232 V=7.0 ACC=20 DEC=20
ARCOF
TIMER T=30
*LAG12
MOVL C00233 V=7.0 ACC=20 DEC=20
MACRO1 MJ#(0) ARGF2
ARCON
MOVL C00234 V=7.0 ACC=20 DEC=20
MOVL C00235 V=7.0 ACC=20 DEC=20
MOVL C00236 V=7.0 ACC=20 DEC=20
MOVL C00237 V=7.0 ACC=20 DEC=20
MOVL C00238 V=7.0 ACC=20 DEC=20
MOVL C00239 V=7.0 ACC=20 DEC=20
MOVL C00240 V=7.0 ACC=20 DEC=20
MOVL C00241 V=7.0 ACC=20 DEC=20
MOVL C00242 V=7.0 ACC=20 DEC=20
MOVL C00243 V=7.0 ACC=20 DEC=20
MOVL C00244 V=7.0 ACC=20 DEC=20
MOVL C00245 V=7.0 ACC=20 DEC=20
MOVL C00246 V=7.0 ACC=20 DEC=20
MOVL C00247 V=7.0 ACC=20 DEC=20
MOVL C00248 V=7.0 ACC=20 DEC=20
MOVL C00249 V=7.0 ACC=20 DEC=20
MOVL C00250 V=7.0 ACC=20 DEC=20
MOVL C00251 V=7.0 ACC=20 DEC=20
MOVL C00252 V=7.0 ACC=20 DEC=20
MOVL C00253 V=7.0 ACC=20 DEC=20
ARCOF
TIMER T=30
*LAG13
MOVL C00254 V=7.0 ACC=20 DEC=20
MACRO1 MJ#(0) ARGF2
ARCON
MOVL C00255 V=7.0 ACC=20 DEC=20
MOVL C00256 V=7.0 ACC=20 DEC=20
MOVL C00257 V=7.0 ACC=20 DEC=20
MOVL C00258 V=7.0 ACC=20 DEC=20
MOVL C00259 V=7.0 ACC=20 DEC=20
MOVL C00260 V=7.0 ACC=20 DEC=20
MOVL C00261 V=7.0 ACC=20 DEC=20
MOVL C00262 V=7.0 ACC=20 DEC=20
MOVL C00263 V=7.0 ACC=20 DEC=20
MOVL C00264 V=7.0 ACC=20 DEC=20
MOVL C00265 V=7.0 ACC=20 DEC=20
MOVL C00266 V=7.0 ACC=20 DEC=20
MOVL C00267 V=7.0 ACC=20 DEC=20
MOVL C00268 V=7.0 ACC=20 DEC=20
MOVL C00269 V=7.0 ACC=20 DEC=20
MOVL C00270 V=7.0 ACC=20 DEC=20
MOVL C00271 V=7.0 ACC=20 DEC=20
MOVL C00272 V=7.0 ACC=20 DEC=20
MOVL C00273 V=7.0 ACC=20 DEC=20
MOVL C00274 V=7.0 ACC=20 DEC=20
ARCOF
TIMER T=30
*LAG14
MOVL C00275 V=7.0 ACC=20 DEC=20
MACRO1 MJ#(0) ARGF2
ARCON
MOVL C00276 V=7.0 ACC=20 DEC=20
MOVL C00277 V=7.0 ACC=20 DEC=20
MOVL C00278 V=7.0 ACC=20 DEC=20
MOVL C00279 V=7.0 ACC=20 DEC=20
MOVL C00280 V=7.0 ACC=20 DEC=20
MOVL C00281 V=7.0 ACC=20 DEC=20
MOVL C00282 V=7.0 ACC=20 DEC=20
MOVL C00283 V=7.0 ACC=20 DEC=20
MOVL C00284 V=7.0 ACC=20 DEC=20
MOVL C00285 V=7.0 ACC=20 DEC=20
MOVL C00286 V=7.0 ACC=20 DEC=20
MOVL C00287 V=7.0 ACC=20 DEC=20
MOVL C00288 V=7.0 ACC=20 DEC=20
MOVL C00289 V=7.0 ACC=20 DEC=20
MOVL C00290 V=7.0 ACC=20 DEC=20
MOVL C00291 V=7.0 ACC=20 DEC=20
MOVL C00292 V=7.0 ACC=20 DEC=20
MOVL C00293 V=7.0 ACC=20 DEC=20
MOVL C00294 V=7.0 ACC=20 DEC=20
MOVL C00295 V=7.0 ACC=20 DEC=20
ARCOF
TIMER T=30
*LAG15
MOVL C00296 V=7.0 ACC=20 DEC=20
MACRO1 MJ#(0) ARGF2
ARCON
MOVL C00297 V=7.0 ACC=20 DEC=20
MOVL C00298 V=7.0 ACC=20 DEC=20
MOVL C00299 V=7.0 ACC=20 DEC=20
MOVL C00300 V=7.0 ACC=20 DEC=20
MOVL C00301 V=7.0 ACC=20 DEC=20
MOVL C00302 V=7.0 ACC=20 DEC=20
MOVL C00303 V=7.0 ACC=20 DEC=20
MOVL C00304 V=7.0 ACC=20 DEC=20
MOVL C00305 V=7.0 ACC=20 DEC=20
MOVL C00306 V=7.0 ACC=20 DEC=20
MOVL C00307 V=7.0 ACC=20 DEC=20
MOVL C00308 V=7.0 ACC=20 DEC=20
MOVL C00309 V=7.0 ACC=20 DEC=20
MOVL C00310 V=7.0 ACC=20 DEC=20
MOVL C00311 V=7.0 ACC=20 DEC=20
MOVL C00312 V=7.0 ACC=20 DEC=20
MOVL C00313 V=7.0 ACC=20 DEC=20
MOVL C00314 V=7.0 ACC=20 DEC=20
MOVL C00315 V=7.0 ACC=20 DEC=20
MOVL C00316 V=7.0 ACC=20 DEC=20
ARCOF
TIMER T=30
MOVL C00317 V=7.0 ACC=20 DEC=20
MOVJ C00318 VJ=0.78
END
